Fanuc KAREL source: STREAM_POS_3.kl

PROGRAM stream_pos_3

%NOLOCKGROUP
%NOPAUSE = ERROR + COMMAND + TPENABLE
%COMMENT = 'CSV -> C1 tag (simple inline)'

VAR
  st     : INTEGER;
  jp     : JOINTPOS;
  cp     : XYZWPR;
  j      : ARRAY[9] OF REAL;
  sock   : FILE;

  t_int  : INTEGER;
  ts_str : STRING[32];
  c_str  : STRING[16];

  s_pre  : STRING[128];
  s_post : STRING[254];
  eol    : STRING[2];
  count  : INTEGER;

  -- Variables for R[25] stop handshake
  r_flag   : BOOLEAN;
  stop_req : INTEGER;
  r_real   : REAL;

ROUTINE rts(val : REAL; digs : INTEGER; decs : INTEGER) : STRING
VAR out : STRING[32];
BEGIN
  CNV_REAL_STR(val, digs, decs, out);
  RETURN(out);
END rts;

BEGIN
  eol = CHR(13) + CHR(10);
  count = 0; -- Initialize the counter

  -- Initialize stop check from R[25]
  GET_REG(25, r_flag, stop_req, r_real, st);

  MSG_CONNECT('C1:', st);
  OPEN FILE sock('RW','C1:');
  IF IO_STATUS(sock) <> 0 THEN
    WRITE('OPEN C1 failed (will retry after first write)'); WRITE(eol);
  ENDIF;

  -- Reordered header (same fields, new order)
  WRITE sock('count,ts_int,ts_str,J1,J2,J3,J4,J5,J6,X,Y,Z,W,P,R'); WRITE sock(eol);

  -- Loop continues while R[25] <> 1
  WHILE (stop_req <> 1) DO
    count = count + 1; -- Increment every loop

    jp = CURJPOS(1, st);
    cp = CURPOS(1, st);
    CNV_JPOS_REL(jp, j, st);

    GET_TIME(t_int);
    CNV_TIME_STR(t_int, ts_str);

    -- Convert the integer count to a string
    CNV_INT_STR(count, 1, 10, c_str);

    -- Start of CSV line: count,
    s_pre  = c_str + ',';

    -- Rest of fields (starts with a comma): J1..J6, X..R
    s_post = ',' +
             rts(j[1],3,6) + ',' + rts(j[2],3,6) + ',' + rts(j[3],3,6) + ',' +
             rts(j[4],3,6) + ',' + rts(j[5],3,6) + ',' + rts(j[6],3,6) + ',' +
             rts(cp.x,3,3) + ',' + rts(cp.y,3,3) + ',' + rts(cp.z,3,3) + ',' +
             rts(cp.w,3,3) + ',' + rts(cp.p,3,3) + ',' + rts(cp.r,3,3);

    -- Write in new order: count, ts_int, ts_str, (then rest)
    WRITE sock(s_pre);
    WRITE sock(t_int);
    WRITE sock(',');
    WRITE sock(ts_str);
    WRITE sock(s_post);
    WRITE sock(eol);

    IF IO_STATUS(sock) <> 0 THEN
      DELAY 200;
      CLOSE FILE sock;
      MSG_DISCO('C1:', st);
      MSG_CONNECT('C1:', st);
      OPEN FILE sock('RW','C1:');

      IF IO_STATUS(sock) = 0 THEN
        -- Reordered header on reconnect too
        WRITE sock('count,ts_int,ts_str,J1,J2,J3,J4,J5,J6,X,Y,Z,W,P,R'); WRITE sock(eol);
      ENDIF;
    ENDIF;

    DELAY 50;

    -- Poll Register 25 every loop iteration
    GET_REG(25, r_flag, stop_req, r_real, st);
  ENDWHILE;

  -- Clean disconnect upon loop exit (R[25] = 1)
  CLOSE FILE sock;
  MSG_DISCO('C1:', st);
END stream_pos_3;
